(* IEC 61131-3 sources: 2026_Projet_YGO_ExcavatriceDragage/TOOLS/TEST_AUTO_CI/MOCKS, 9 files *)

(* ---- DEVICE_STATE.st ---- *)
(* =======================================================================
   📊 Type CODESYS système pour tests STruCpp
   ======================================================================= *)
TYPE DEVICE_STATE :
(
    UNKNOWN             := 0,
    STOPPED             := 1,
    CONFIG_ERROR        := 2,
    BUS_ERROR           := 3,
    DISABLED            := 4,
    INITIALIZING        := 5,
    RESET_ORIGIN        := 6,
    RESET_COMMUNICATION := 7,
    RESET_APPLICATION   := 8,
    RUNNING             := 9,
    LOGGER_ERROR        := 10
);
END_TYPE

(* ---- MOCK_GVL_IHM.st ---- *)
(* =======================================================================
   🧪 MOCK_GVL_IHM — Miroir TESTABLE de la GVL_IHM (harnais CI uniquement)
   ───────────────────────────────────────────────────────────────
   🎯 Pourquoi ce fichier existe (T371) :
      STruCpp v0.6.2 ne supporte PAS le namespace GVL de CODESYS. Une GVL
      `VAR_GLOBAL` déclare ses membres comme des variables GLOBALES PLATES :
      `GVL_IHM.Modes.Cmd.X` n'est donc pas résoluble, alors que c'est
      exactement ce que fait le code de production (CODESYS, où le nom de la
      GVL EST un espace de noms).
      Sonde compilateur (2026-09-21) : `VAR_GLOBAL Foo:INT;` + `GVL_T.Foo`
      -> "error: Undeclared variable 'GVL_T'" ; accès direct `Foo` -> OK ;
      `GVL_T` déclaré comme VARIABLE d'un STRUCT miroir -> OK.

   🔧 Principe : `GVL_IHM` est déclarée ici comme une VARIABLE GLOBALE d'un
      STRUCT MIROIR dont les membres sont la TRANSCRIPTION EXACTE de la liste
      de membres de `CODE/J_SUPERVISION/GVL_IHM.st`. Le code de production
      (`GVL_IHM.<membre>`) devient alors résoluble à l'identique.

   ⚠️ FICHIER DE TEST — JAMAIS compilé dans CODESYS, JAMAIS importé :
      il n'est référencé que par l'entrée `FB_TroubleshootingView` de
      `TOOLS/TEST_AUTO_CI/scripts/config/registry.yaml`.
   ⚠️ DETTE DÉCLARÉE : ce miroir peut dériver si `GVL_IHM.st` change. Une
      dérive produit une ERREUR DE COMPILATION du harnais (bruit), jamais un
      faux résultat silencieux. Toute évolution de `GVL_IHM.st` doit être
      répercutée ici.
   📄 Source de vérité transcrite : CODE/J_SUPERVISION/GVL_IHM.st:8-24
   ======================================================================= *)

TYPE ST_MockGvlIHM :
STRUCT
    M1TreuilRetenue    : ST_WinchHMI;               (* GVL_IHM.st:8  *)
    M2TreuilBenne      : ST_WinchBenneHMI;          (* GVL_IHM.st:9  — porte Bucket *)
    M1M2Sync           : ST_SyncHMI;                (* GVL_IHM.st:10 *)
    JOY1Joystick       : ST_JoystickHMI;            (* GVL_IHM.st:11 *)
    Modes              : ST_ModesHMI;               (* GVL_IHM.st:12 *)
    Emergency          : ST_EmergencyHMI;           (* GVL_IHM.st:13 *)
    M3Translation      : ST_TranslationHMI;         (* GVL_IHM.st:14 *)
    CycleSemiAuto      : ST_CycleHMI;               (* GVL_IHM.st:15 *)
    CycleMachineHoming : ST_CycleMachineHomingHMI;  (* GVL_IHM.st:16 *)
    Banner             : ST_HmiBanner;              (* GVL_IHM.st:17 *)
    Network            : ST_NetworkDiagHMI;         (* GVL_IHM.st:18 *)
    Commun             : ST_CommunHMI;              (* GVL_IHM.st:19 *)
    LocalIHM           : ST_LocalIHM;               (* GVL_IHM.st:20 *)
    IoHw               : ST_IoHw;                   (* GVL_IHM.st:21 *)
    HmiInitDone        : BOOL;                      (* GVL_IHM.st:22 *)
    Permits            : ST_PermitVisibilityHMI;    (* GVL_IHM.st:23 *)
    MaintenanceN2      : ST_MaintenanceN2HMI;       (* GVL_IHM.st:24 *)
END_STRUCT
END_TYPE

VAR_GLOBAL
    GVL_IHM : ST_MockGvlIHM;   // Miroir testable de la GVL de production (voir bandeau)
END_VAR

(* ---- MOCK_GVL_Troubleshooting.st ---- *)
(* =======================================================================
   🧪 MOCK_GVL_Troubleshooting — Miroir TESTABLE de la GVL_Troubleshooting
   ───────────────────────────────────────────────────────────────
   🎯 Pourquoi ce fichier existe (T371) : voir le bandeau détaillé de
      `TOOLS/TEST_AUTO_CI/MOCKS/MOCK_GVL_IHM.st` (même cause, même patron).
      En résumé : STruCpp v0.6.2 ne supporte pas le namespace GVL CODESYS ;
      `GVL_Troubleshooting.N_MotionM1.Step8_OutputInterlockOk` (écrit 469 fois
      par `FB_TroubleshootingView.st`) n'est résoluble que si `GVL_Troubleshooting`
      existe comme VARIABLE GLOBALE d'un STRUCT miroir — patron prouvé par sonde
      compilateur le 2026-09-21.

   ⚠️ FICHIER DE TEST — JAMAIS compilé dans CODESYS, JAMAIS importé :
      référencé uniquement par l'entrée `FB_TroubleshootingView` du registry CI.
   ⚠️ DETTE DÉCLARÉE : dérive possible si `GVL_Troubleshooting.st` change ->
      erreur de compilation du harnais (bruit), jamais un faux résultat silencieux.
   📄 Source de vérité transcrite : CODE/J_SUPERVISION/GVL_Troubleshooting.st
      (bloc VAR_GLOBAL, membres dans l'ordre du fichier source)
   ======================================================================= *)

TYPE ST_MockGvlTroubleshooting :
STRUCT
    A_ContexteMachineGlobal  : ST_ChainContextGlobal;   (* 0.  Contexte Global Machine *)
    B_Inputs                 : ST_HardwareImage;        (* 1.  Image complète des entrées *)
    C_Safety                 : ST_SafetyChecklist;      (* 2.  Chaîne de sécurité & réarmement AU *)
    D_Joystick               : ST_JoystickChecklist;    (* 3.  Bus CANopen & homme-mort joystick *)
    E_HomingM1               : ST_HomingChecklist;      (* 4.  Homing M1 *)
    F_HomingM2               : ST_HomingChecklist;      (* 5.  Homing M2 *)
    G_CycleSemiAuto          : ST_ChainCycleSemiAuto;   (* 6.  Séquenceur de cycle semi-auto *)
    H_LevageSynchroniseM1M2  : ST_ChainWinchSync;       (* 7.  Levage synchronisé M1+M2 *)
    I_LevageUnitaireM1       : ST_ChainWinch;           (* 8.  Levage unitaire M1 *)
    J_LevageUnitaireM2       : ST_ChainWinch;           (* 9.  Levage unitaire M2 *)
    K_BenneOuvertureFermeture: ST_ChainBucket;          (* 10. Ouverture / fermeture benne *)
    L_TranslationPontM3      : ST_ChainTranslation;     (* 11. Translation pont M3 *)
    N_MotionM1               : ST_MotionChecklist;      (* 13. Diagnostic mouvement M1 *)
    O_MotionM2               : ST_MotionChecklist;      (* 14. Diagnostic mouvement M2 *)
    P_MotionM3               : ST_MotionChecklist;      (* 15. Diagnostic mouvement M3 *)
    Q_TraceWinchM1           : ST_TraceWinch;           (* 16. Trace blocage M1 *)
    R_TraceWinchM2           : ST_TraceWinch;           (* 17. Trace blocage M2 *)
    S_TraceTranslation       : ST_TraceTranslation;     (* 18. Trace blocage M3 *)
    T_Permits                : ST_PermitVisibilityHMI;  (* Vue unique des permis *)
END_STRUCT
END_TYPE

VAR_GLOBAL
    GVL_Troubleshooting : ST_MockGvlTroubleshooting;   // Miroir testable de la GVL de production
END_VAR

(* ---- ST_fbJoystick_Cfg.st ---- *)
(* =======================================================================
   🧪 ST_fbJoystick_Cfg — Maquette STruCpp pour FB_SimBench
   -----------------------------------------------------------------------
   🎯 Rôle : satisfaire le champ ST_JoystickHMI.Cfg sans exercer FB_Joystick.
   📄 Portée : harnais STruCpp uniquement; le type production reste inchangé.
   ======================================================================= *)
TYPE ST_fbJoystick_Cfg :
STRUCT
END_STRUCT
END_TYPE

(* ---- ST_fbSim_Translation_ExtLink_Echo.st ---- *)
(* Test-only mirror of the retired external-M3 link payload.
   Production code no longer ships the OpenModelica link; FB_SimBench CI still
   requires its interface because MOCK_FB_Sim_Translation_ExtLink exposes it. *)
TYPE ST_fbSim_Translation_ExtLink_Echo :
STRUCT
    Mode                    : E_Mode;
    FBState                 : E_State;
    AxisBlockReason         : E_TranslationTraceBlockReason;
    MaintenanceTargetEnable : BOOL;
    MaintenanceZoneAccess   : BOOL;
    SafeStop                : BOOL;
    PowerCutOff             : BOOL;
    LimitSwitchTremie       : BOOL;
    LimitSwitchMaintenance  : BOOL;
    PositionReached         : BOOL;
    ActiveTremie            : BOOL;
    ActiveMaintenance       : BOOL;
    AtTremie                : BOOL;
    AtPV                    : BOOL;
    AtP2                    : BOOL;
    AtP1                    : BOOL;
    AtMaintenance           : BOOL;
    SensorWordIncoherent    : BOOL;
    EstimatedPos_M          : REAL;
    SafetyErrorId           : WORD;
END_STRUCT
END_TYPE

(* ---- FB_TestHarnessT417_M3.st ---- *)
(* T417 D2 — boucle fermee de preuve, composants de production composes dans l'ordre PRG02→PRG03/05→PRG06.
   Le cycle utilise ses entrees publiques. StepForceTgt ne sert qu'a fixer le point de depart AX14;
   les gestes, les transitions AX15A/B/C/18/2 et les demandes M3 restent emis par les vrais FB.
   M1/M2, benne, mode arbitre, IHM, reseaux et AU sont des faits de banc declares, pas couverts ici. *)
FUNCTION_BLOCK PUBLIC FB_TestHarnessT417_M3
VAR_INPUT
    Enable                  : BOOL;
    StepForceTgt            : INT := -1;
    JoystickLeft            : BOOL;
    JoystickRight           : BOOL;
    JoystickPush            : BOOL;
    JoystickPull            : BOOL;
    RepositionRequest       : BOOL;
    BenneDone               : BOOL;
    BenneIsOpen             : BOOL;
    SimM3Slope_Mps2         : REAL;
END_VAR
VAR_IN_OUT
    RawPosM1                : UDINT;
    RawPosM2                : UDINT;
END_VAR
VAR_OUTPUT
    CycleStep               : E_AutoCycleStep;
    CycleError              : BOOL;
    CycleReqStart            : BOOL;
    CyclePositionTgt          : INT;
    ArbitrationReqTremie      : BOOL;
    ArbitrationReqMaintenance : BOOL;
    ArbitrationRunRequest     : BOOL;
    TranslationSafetyError  : BOOL;
    TranslationMotionError  : BOOL;
    FinalInterlockError     : BOOL;
    M3ReqTremie              : BOOL;
    M3ReqMaintenance         : BOOL;
    M3DriveControlWord       : WORD;
    M3DriveFreqCmd_Hz        : REAL;
    M3DriveActualFreq_Hz     : REAL;
    M3BrakeReleaseRequest    : BOOL;
    M3BrakeFinalCmd          : BOOL;
    M3BrakeContactOpen       : BOOL;
    M3SensorsWord            : BYTE;
    M3AtTremie               : BOOL;
    M3AtP1                   : BOOL;
    M3PositionTrue_M         : REAL;
    M3PositionEstimated_M    : REAL;
    M3PositionError_M        : REAL;
    M3OvershootLast_M        : REAL;
    M3OvershootSensorId      : INT;
    P1ArrivalCaptured        : BOOL;
    P1ArrivalPosition_M       : REAL;
    P1ArrivalSensorsWord      : BYTE;
    P1ArrivalDriveControlWord : WORD;
    P1ArrivalFrequency_Hz     : REAL;
    P1ArrivalBrakeOpen        : BOOL;
    M3CartFree               : BOOL;
    M3FreeRollLast_M         : REAL;
END_VAR
VAR
    instCycle                : FB_CycleSemiAuto;
    instArbitration          : FB_TranslationCmdArbitrationM3;
    instSafety               : FB_Safety_Translation;
    instTranslation          : FB_Translation;
    instOutputInterlock      : FB_TranslationOutputInterlock;
    instPositionDecoder      : FB_Translation_PositionDecoder;
    instPositionEstimator    : FB_Translation_PositionEstimator;
    instSimBench             : FB_SimBench;
    TranslationCfg           : ST_fbTranslation_Cfg;
    Joystick                 : ST_AcquisitionJoystickQualified;
    ModesAuth                : ST_Modes_Autorisations;
    CycleTranslationRequest  : ST_ProgramTranslationRequest;
    ArbitrationIHM           : ST_fbTranslationCmdArbitration_IHM;
    ArbitrationContext       : ST_fbTranslationCmdArbitration_Context;
    ArbitrationCfg           : ST_fbTranslationCmdArbitration_Cfg;
    TargetCodeSel            : INT;
    SensorsWordPrev          : BYTE;
    SensorsWordChanged       : BOOL;
    PositionSensorTarget     : BOOL;
    AtTremieStable           : BOOL;
    AtPVStable               : BOOL;
    AtP2Stable               : BOOL;
    AtP1Stable               : BOOL;
    AtMaintenanceStable      : BOOL;
    AtPositionBootRestored   : BOOL;
    BootSensorsStable        : TON;
    SimReqTremieN1           : BOOL;
    SimReqMaintenanceN1      : BOOL;
    SimSpeedPctN1            : REAL;
    SimBrakeCmdN1            : BOOL;
    M3HeightInterlockOk      : BOOL;
    PermitTremie             : BOOL;
    PermitMaintenance        : BOOL;
    P1ArrivalCapturedLocal    : BOOL;
END_VAR

IF NOT Enable THEN
    CycleStep := E_AutoCycleStep.AX0_REPOS;
    RETURN;
END_IF;

(* La simulation est PRG02 : elle consomme les sorties finales mémorisées du scan N-1. *)
instSimBench(
    Enable := TRUE,
    OperatorSourceActive := TRUE,
    M3_ReqTremie := SimReqTremieN1,
    M3_ReqMaintenance := SimReqMaintenanceN1,
    M3_SpeedCmd_Pct := SimSpeedPctN1,
    M3_PosTremie_M := 0.0,
    M3_PosPV_M := 1.5,
    M3_PosP2_M := 3.5,
    M3_PosP1_M := 5.0,
    M3_PosMaintenance_M := 10.0,
    M3_OdometryGain := 0.02,
    M3_EstimatedPos_M := instPositionEstimator.PositionEstimatedM,
    M3_BrakeCmd := SimBrakeCmdN1,
    PowerKeepAlive_A := TRUE,
    PowerKeepAlive_B := TRUE,
    SimChainOkBit := TRUE,
    SimPhaseRotationOkBit := TRUE,
    SimM3SpeedFactor := 1.0,
    SimM3SensorIntermittenceActive := FALSE,
    SimM3SensorCamDropoutActive := FALSE,
    SimM3BrakePhysicalActive := TRUE,
    SimM3CartFreeActive := TRUE,
    SimM3LoadMassRatio := 0.5,
    SimM3RollingFriction_Mps2 := 0.1,
    SimM3Slope_Mps2 := SimM3Slope_Mps2,
    RawPosM1 := RawPosM1,
    RawPosM2 := RawPosM2
);

instPositionDecoder(
    SensorTremie := instSimBench.Translation.M3_PosTremie_DI,
    SensorPV := instSimBench.Translation.M3_PosPV_DI,
    SensorP2 := instSimBench.Translation.M3_PosPVP2_DI,
    SensorP1 := instSimBench.Translation.M3_PosP1_DI,
    SensorMaintenance := instSimBench.Translation.M3_PosMaintenance_DI
);

instPositionEstimator(
    Enable := TRUE,
    Reset := FALSE,
    DriveActualFreqHz := UINT_TO_REAL(instSimBench.Translation.M3_ActualFrequencyHz) / 100.0,
    ReqTremie := SimReqTremieN1,
    ReqMaintenance := SimReqMaintenanceN1,
    SensorMaintenance := instPositionDecoder.TranslationPosMaintenance,
    SensorP1 := instPositionDecoder.TranslationPosP1,
    SensorP2 := instPositionDecoder.TranslationPosP2,
    SensorPV := instPositionDecoder.TranslationPosPV,
    SensorTremie := instPositionDecoder.TranslationPosTremie,
    PosMaintenanceM := 10.0,
    PosP1M := 5.0,
    PosP2M := 3.5,
    PosPVM := 1.5,
    PosTremieM := 0.0,
    GainMetersPerHzSec := 0.02,
    PersistedPositionM := 0.0,
    PersistedInitialized := FALSE
);

SensorsWordChanged := instPositionDecoder.SensorsWord <> SensorsWordPrev;
BootSensorsStable(IN := NOT SimReqTremieN1 AND NOT SimReqMaintenanceN1, PT := T#500ms);
IF NOT AtPositionBootRestored AND BootSensorsStable.Q THEN
    CASE instPositionDecoder.SensorsWord OF
        2#11111: AtTremieStable := instPositionDecoder.TranslationPosTremie;
        2#01111: AtPVStable := instPositionDecoder.TranslationPosPV;
        2#00111: AtP2Stable := instPositionDecoder.TranslationPosP2;
        2#00011: AtP1Stable := instPositionDecoder.TranslationPosP1;
        2#00000: AtMaintenanceStable := instPositionDecoder.TranslationPosMaintenance;
    END_CASE;
    AtPositionBootRestored := TRUE;
ELSIF AtPositionBootRestored THEN
    IF instPositionDecoder.TranslationAtTremie THEN
        AtTremieStable := TRUE; AtPVStable := FALSE; AtP2Stable := FALSE; AtP1Stable := FALSE; AtMaintenanceStable := FALSE;
    ELSIF instPositionDecoder.TranslationAtPV THEN
        AtPVStable := TRUE; AtTremieStable := FALSE; AtP2Stable := FALSE; AtP1Stable := FALSE; AtMaintenanceStable := FALSE;
    ELSIF instPositionDecoder.TranslationAtP2 THEN
        AtP2Stable := TRUE; AtTremieStable := FALSE; AtPVStable := FALSE; AtP1Stable := FALSE; AtMaintenanceStable := FALSE;
    ELSIF instPositionDecoder.TranslationAtP1 THEN
        AtP1Stable := TRUE; AtTremieStable := FALSE; AtPVStable := FALSE; AtP2Stable := FALSE; AtMaintenanceStable := FALSE;
    ELSIF instPositionDecoder.TranslationAtMaintenance THEN
        AtMaintenanceStable := TRUE; AtTremieStable := FALSE; AtPVStable := FALSE; AtP2Stable := FALSE; AtP1Stable := FALSE;
    ELSIF SensorsWordChanged THEN
        AtPVStable := FALSE; AtP2Stable := FALSE; AtP1Stable := FALSE;
    END_IF;
    IF SimReqMaintenanceN1 THEN AtTremieStable := FALSE; END_IF;
    IF SimReqTremieN1 THEN AtMaintenanceStable := FALSE; END_IF;
END_IF;
SensorsWordPrev := instPositionDecoder.SensorsWord;

Joystick.AxisX.Enable := TRUE;
Joystick.AxisX.StartStop := JoystickLeft OR JoystickRight;
Joystick.AxisX.DirectionPositive := JoystickLeft;
Joystick.AxisX.DirectionNegative := JoystickRight;
Joystick.AxisX.AtNeutral := NOT JoystickLeft AND NOT JoystickRight;
Joystick.AxisX.Direction := SEL(JoystickLeft, SEL(JoystickRight, 0, -1), 1);
Joystick.AxisX.SpeedTgt := 100.0;
Joystick.AxisY.Enable := TRUE;
Joystick.AxisY.StartStop := JoystickPush OR JoystickPull;
Joystick.AxisY.DirectionPositive := JoystickPush;
Joystick.AxisY.DirectionNegative := JoystickPull;
Joystick.AxisY.AtNeutral := NOT JoystickPush AND NOT JoystickPull;
Joystick.AxisY.Direction := SEL(JoystickPush, SEL(JoystickPull, 0, -1), 1);
Joystick.AxisY.SpeedTgt := 100.0;
Joystick.DeadmanArmed := TRUE;
Joystick.AtNeutralXY := Joystick.AxisX.AtNeutral AND Joystick.AxisY.AtNeutral;
Joystick.Ready := TRUE;
ModesAuth.Mode := E_Mode.SEMI_AUTO;
ModesAuth.MaintenanceM3TargetEnable := FALSE;
M3HeightInterlockOk := TRUE; (* entree de banc declaree : M1/M2 au-dessus du seuil de PRG05 *)

instCycle(
    Enable := TRUE,
    PowerContactorEngaged := TRUE,
    EncoderFaultPresent := FALSE,
    Mode := E_Mode.SEMI_AUTO,
    JoystickDeflected := JoystickLeft OR JoystickRight OR JoystickPush OR JoystickPull,
    JoystickPush := JoystickPush,
    JoystickPull := JoystickPull,
    JoystickRight := JoystickRight,
    JoystickLeft := JoystickLeft,
    DeadmanArmed := TRUE,
    HeartbeatIhmOk := TRUE,
    SelTarget := 0,
    SetDepthM := -5.0,
    DepthStopMode := E_CycleDepthStopMode.KOBOLD_ONLY,
    WinchSyncError := FALSE,
    WinchSyncDeltaM := 0.0,
    M1_CablePosM := 5.0,
    M2_CablePosM := 5.0,
    M1_MeasuredSpeedMps := 0.0,
    M2_MeasuredSpeedMps := 0.0,
    M1_SpeedValid := TRUE,
    M2_SpeedValid := TRUE,
    M1_ContactorsReleased := TRUE,
    M2_ContactorsReleased := TRUE,
    M1_BrakeApplied := TRUE,
    M2_BrakeApplied := TRUE,
    SpeedMismatchThresholdMps := 0.0,
    SpeedMismatchTimeout := T#0ms,
    M1TopLimitReached := TRUE,
    M2TopLimitReached := TRUE,
    Translation_At_P1 := AtP1Stable,
    Translation_At_Tremie := AtTremieStable,
    Translation_At_Maintenance := AtMaintenanceStable,
    Translation_PosP1 := instPositionDecoder.TranslationPosP1,
    Translation_PosMaintenance := instPositionDecoder.TranslationPosMaintenance,
    Translation_Busy := ABS(instTranslation.RequestedDriveFreqHz) > 0.1,
    Translation_Done := instTranslation.TargetReached,
    Benne_Done := BenneDone,
    Benne_CloseReached := NOT BenneIsOpen,
    Benne_IsOpen := BenneIsOpen,
    Benne_IsClosed := NOT BenneIsOpen,
    Benne_IsRoughlyClosed := NOT BenneIsOpen,
    M1FinalAscentStartReady := TRUE,
    HomedM1 := TRUE,
    HomedM2 := TRUE,
    InitPositionOk := TRUE,
    WinchesAtTopWindow := TRUE,
    CfgDrainTime := T#0ms,
    RepositionRequest := RepositionRequest,
    StepForceTgt := StepForceTgt
);
CycleStep := instCycle.CycleStep;
CycleError := instCycle.Fault.Error;
CycleTranslationRequest := instCycle.TranslationCmd;
CycleReqStart := CycleTranslationRequest.ReqStart;
CyclePositionTgt := CycleTranslationRequest.PositionTgt;

ArbitrationContext.HeightInterlockOk := M3HeightInterlockOk;
ArbitrationCfg.MaxFreq_Hz := 50.0;
instArbitration(
    Enable := TRUE,
    Joystick := Joystick,
    Auth := ModesAuth,
    ReqTranslation := CycleTranslationRequest,
    IHM := ArbitrationIHM,
    TglJoystickMaster := FALSE,
    Context := ArbitrationContext,
    Cfg := ArbitrationCfg
);
ArbitrationReqTremie := instArbitration.ReqTremie;
ArbitrationReqMaintenance := instArbitration.ReqMaintenance;
ArbitrationRunRequest := instArbitration.RunRequest;
(* Le selecteur de cible est consommable au scan courant : retenir la derniere valeur non nulle. *)
IF instArbitration.SelTarget >= 1 AND instArbitration.SelTarget <= 4 THEN
    TargetCodeSel := instArbitration.SelTarget;
END_IF;
IF instArbitration.SelTarget = 0 THEN
    IF instArbitration.ReqTremie THEN
        TargetCodeSel := 1;
    ELSIF instArbitration.ReqMaintenance THEN
        TargetCodeSel := SEL(ModesAuth.MaintenanceM3TargetEnable, 3, 4);
    END_IF;
END_IF;
PositionSensorTarget := FALSE;
CASE TargetCodeSel OF
    1: PositionSensorTarget := AtTremieStable;
    2: PositionSensorTarget := AtP2Stable;
    3: PositionSensorTarget := AtP1Stable;
    4: PositionSensorTarget := AtMaintenanceStable;
END_CASE;

instSafety(
    Enable := TRUE,
    Reset := FALSE,
    PowerContactorEngaged := TRUE,
    Mode := E_Mode.SEMI_AUTO,
    JoystickOnline := TRUE,
    JoystickOperational := TRUE,
    HeartbeatIhmOk := TRUE,
    PhaseRotationOk := TRUE,
    BrakeThermalFeedback := FALSE,
    DriveOnline := TRUE,
    DriveOperational := TRUE,
    DriveStatusWord := instSimBench.Translation.M3_StatusWord,
    DriveActualFreqHz := UINT_TO_REAL(instSimBench.Translation.M3_ActualFrequencyHz) / 100.0,
    BrakeFeedback := instSimBench.Translation.M3_BrakeIsOpen_DI,
    BrakeCmd := instTranslation.BrakeReleaseRequest,
    RunRequest := instArbitration.RunRequest,
    ReqTremie := instArbitration.ReqTremie,
    ReqMaintenance := instArbitration.ReqMaintenance,
    LimitSwitchTremie := instPositionDecoder.LimitSwitchTremie,
    LimitSwitchMaintenance := instPositionDecoder.LimitSwitchMaintenance,
    SensorWordIncoherent := instPositionDecoder.Incoherent
);
PermitTremie := instSafety.TremieLimitClear AND NOT instSafety.SafeStop AND NOT instSafety.PowerCutOff;
PermitMaintenance := instSafety.MaintenanceLimitClear AND NOT instSafety.SafeStop AND NOT instSafety.PowerCutOff;

TranslationCfg.CfgRampAccelRate := 40.0;
TranslationCfg.CfgRampDecelNormalRate := 50.0;
TranslationCfg.CfgRampDecelFastRate := 100.0;
TranslationCfg.DriveFreqScaleMaxHz := 50.0;
TranslationCfg.ApproachSpeedTremieHz := 20.0;
TranslationCfg.ApproachSpeedMaintenanceHz := 20.0;
TranslationCfg.ApproachSpeedP1Hz := 20.0;
instTranslation(
    Enable := TRUE,
    Reset := FALSE,
    PowerContactorEngaged := TRUE,
    Mode := E_Mode.SEMI_AUTO,
    RunRequest := instArbitration.RunRequest,
    SafeStop := instSafety.SafeStop,
    ReqTremie := instArbitration.ReqTremie,
    ReqMaintenance := instArbitration.ReqMaintenance,
    SpeedTgt_Pct := instArbitration.SpeedPct,
    PositionSensorTarget := PositionSensorTarget,
    SlowdownSensorTremie := instPositionDecoder.TranslationPosPV,
    SlowdownSensorMaintenance := instPositionDecoder.TranslationPosP1,
    SlowdownSensorP1 := (NOT instPositionDecoder.TranslationPosP2) AND instPositionDecoder.TranslationPosP1,
    LimitSwitchTremie := instPositionDecoder.LimitSwitchTremie,
    LimitSwitchMaintenance := instPositionDecoder.LimitSwitchMaintenance,
    EffectivePermitM3_Tremie := PermitTremie,
    EffectivePermitM3_Maintenance := PermitMaintenance,
    DriveStatusWord := instSimBench.Translation.M3_StatusWord,
    DriveActualFreqHz := UINT_TO_REAL(instSimBench.Translation.M3_ActualFrequencyHz) / 100.0,
    BrakeFeedback := instSimBench.Translation.M3_BrakeIsOpen_DI,
    Cfg := TranslationCfg
);

instOutputInterlock(
    Enable := TRUE,
    Reset := FALSE,
    SafeStop := instSafety.SafeStop,
    PowerContactorEngaged := TRUE,
    EffectivePermitM3_Tremie := PermitTremie,
    EffectivePermitM3_Maintenance := PermitMaintenance,
    BrakeReleaseRequest := instTranslation.BrakeReleaseRequest,
    BrakeCommandOpenConfirmed := instTranslation.BrakeCommandOpenConfirmed,
    RequestedDriveControlWord := instTranslation.RequestedDriveControlWord,
    RequestedDriveFreqHz := instTranslation.RequestedDriveFreqHz
);

SimReqTremieN1 := instOutputInterlock.DriveControlWord = 1;
SimReqMaintenanceN1 := instOutputInterlock.DriveControlWord = 2;
SimSpeedPctN1 := (instOutputInterlock.DriveFreqCmd_Hz / 50.0) * 100.0;
SimBrakeCmdN1 := instOutputInterlock.BrakeCmd;

TranslationSafetyError := instSafety.Fault.Error;
TranslationMotionError := instTranslation.Fault.Error;
FinalInterlockError := instOutputInterlock.Fault.Error;
M3ReqTremie := SimReqTremieN1;
M3ReqMaintenance := SimReqMaintenanceN1;
M3DriveControlWord := instOutputInterlock.DriveControlWord;
M3DriveFreqCmd_Hz := instOutputInterlock.DriveFreqCmd_Hz;
M3DriveActualFreq_Hz := UINT_TO_REAL(instSimBench.Translation.M3_ActualFrequencyHz) / 100.0;
M3BrakeReleaseRequest := instTranslation.BrakeReleaseRequest;
M3BrakeFinalCmd := instOutputInterlock.BrakeCmd;
M3BrakeContactOpen := instSimBench.Translation.M3_BrakeIsOpen_DI;
M3SensorsWord := instPositionDecoder.SensorsWord;
M3AtTremie := AtTremieStable;
M3AtP1 := AtP1Stable;
M3PositionTrue_M := instSimBench.M3ObsPositionTrue_M;
M3PositionEstimated_M := instPositionEstimator.PositionEstimatedM;
M3PositionError_M := instSimBench.M3ObsPositionError_M;
M3OvershootLast_M := instSimBench.M3ObsOvershootLast_M;
M3OvershootSensorId := instSimBench.M3ObsOvershootSensorId;
IF (CycleStep = E_AutoCycleStep.AX18_DONE_SYNC) THEN
    P1ArrivalCapturedLocal := FALSE;
END_IF;
IF (CycleStep = E_AutoCycleStep.AX2_TRANSLATE_P1) AND AtP1Stable AND NOT P1ArrivalCapturedLocal THEN
    P1ArrivalCapturedLocal := TRUE;
    P1ArrivalCaptured := TRUE;
    P1ArrivalPosition_M := M3PositionTrue_M;
    P1ArrivalSensorsWord := M3SensorsWord;
    P1ArrivalDriveControlWord := M3DriveControlWord;
    P1ArrivalFrequency_Hz := M3DriveActualFreq_Hz;
    P1ArrivalBrakeOpen := M3BrakeContactOpen;
END_IF;
M3CartFree := instSimBench.M3ObsCartFree;
M3FreeRollLast_M := instSimBench.M3ObsFreeRollLast_M;
END_FUNCTION_BLOCK

(* ---- FB_TestLoopTranslation.st ---- *)
(* Harnais de test T417 : boucle fermee FB_Translation REEL (non modifie) + decodeur + FB_Sim_Translation.
   Un appel = un scan. Reproduit le cablage de PRG_05 (decodeur, ralentissements d approche, FdC bistable P1
   quand Maintenance est interdite, permis, jeton d arrivee P1). Non reproduit : FB_TranslationOutputInterlock
   (traite en transparent) et FB_Safety_Translation. Cible P1. Jamais compile dans le programme CODESYS. *)
FUNCTION_BLOCK FB_TestLoopTranslation
VAR_INPUT
    HoldRequest : BOOL;
END_VAR
VAR_OUTPUT
    Phase : INT;
    Overshoot_M : REAL;
    FreqAtCross_Hz : REAL;
    MaxCmdAfter_Hz : REAL;
    PositionTrue_M : REAL;
    CtrlWord : WORD;
    FreqReq_Hz : REAL;
    ActualFreq_Hz : REAL;
    AtP1Token : BOOL;
    SensorsWord : BYTE;
END_VAR
VAR
    tr : FB_Translation;
    sim : FB_Sim_Translation;
    dec : FB_Translation_PositionDecoder;
    cfg : ST_fbTranslation_Cfg;
    Initialized : BOOL;
    reqTremie : BOOL;
    reqMaint : BOOL;
    limTremieStable : BOOL;
    limMaintStable : BOOL;
    limMaintEff : BOOL;
    atP1 : BOOL;
    wordPrev : BYTE;
    wordChanged : BOOL;
    stopCount : INT;
    maxPos_M : REAL;
    crossed : BOOL;
END_VAR

IF NOT Initialized THEN
    Initialized := TRUE;
    cfg.CfgRampAccelRate := 40.0;
    cfg.CfgRampDecelNormalRate := 50.0;
    cfg.CfgRampDecelFastRate := 100.0;
    cfg.DriveFreqScaleMaxHz := 50.0;
    cfg.ApproachSpeedTremieHz := 20.0;
    cfg.ApproachSpeedMaintenanceHz := 20.0;
    cfg.ApproachSpeedP1Hz := 20.0;
    Phase := 0;
    reqTremie := TRUE;
END_IF;

dec(SensorTremie := sim.PosTremie, SensorPV := sim.PosPV, SensorP2 := sim.PosP2,
    SensorP1 := sim.PosP1, SensorMaintenance := sim.PosMaintenance);
limMaintEff := (NOT dec.TranslationPosP1) AND dec.TranslationPosMaintenance;
IF dec.LimitSwitchTremie THEN
    limTremieStable := TRUE;
ELSIF reqMaint THEN
    limTremieStable := FALSE;
END_IF;
IF limMaintEff THEN
    limMaintStable := TRUE;
ELSIF reqTremie THEN
    limMaintStable := FALSE;
END_IF;
wordChanged := (dec.SensorsWord <> wordPrev);
wordPrev := dec.SensorsWord;
IF dec.TranslationAtP1 THEN
    atP1 := TRUE;
ELSIF dec.TranslationAtP2 OR dec.TranslationAtPV OR dec.TranslationAtTremie OR dec.TranslationAtMaintenance OR wordChanged THEN
    atP1 := FALSE;
END_IF;

tr(Enable := TRUE, Reset := FALSE, PowerContactorEngaged := TRUE, RunRequest := TRUE, SafeStop := FALSE,
   ReqTremie := reqTremie, ReqMaintenance := reqMaint, SpeedTgt_Pct := 100.0,
   PositionSensorTarget := atP1 AND reqMaint,
   SlowdownSensorTremie := dec.TranslationPosPV,
   SlowdownSensorMaintenance := (NOT dec.TranslationPosP1) AND dec.TranslationPosMaintenance,
   SlowdownSensorP1 := (NOT dec.TranslationPosP2) AND dec.TranslationPosP1,
   LimitSwitchTremie := limTremieStable, LimitSwitchMaintenance := limMaintStable,
   EffectivePermitM3_Tremie := NOT limTremieStable, EffectivePermitM3_Maintenance := NOT limMaintStable,
   DriveStatusWord := 0, DriveActualFreqHz := sim.ActualFrequency_Hz,
   BrakeFeedback := sim.BrakeContactOpen, Cfg := cfg);
sim(Enable := TRUE,
    ReqTremie := (tr.RequestedDriveControlWord = 1), ReqMaintenance := (tr.RequestedDriveControlWord = 2),
    SpeedTgt_Pct := LIMIT(0.0, tr.RequestedDriveFreqHz / 50.0 * 100.0, 100.0),
    BrakeReleaseCmd := tr.BrakeReleaseRequest,
    LoadFrequencyDroopGain_Hz := 0.0, LoadReactionGain_Mps2 := 0.0);
PositionTrue_M := sim.PositionTrue_M;
CtrlWord := tr.RequestedDriveControlWord;
FreqReq_Hz := tr.RequestedDriveFreqHz;
ActualFreq_Hz := sim.ActualFrequency_Hz;
AtP1Token := atP1;
SensorsWord := dec.SensorsWord;

CASE Phase OF
    0:  (* jambe Tremie jusqu a 6 m : vitesse pleine atteinte hors zone d approche *)
        IF sim.PositionTrue_M < 6.0 THEN
            reqTremie := FALSE;
            Phase := 1;
            stopCount := 0;
        END_IF;
    1:  (* arret complet, frein ferme *)
        IF (sim.ActualFrequency_Hz < 0.5) AND (NOT sim.BrakeMechanicallyOpen) THEN
            stopCount := stopCount + 1;
        ELSE
            stopCount := 0;
        END_IF;
        IF stopCount > 30 THEN
            reqMaint := TRUE;
            Phase := 2;
        END_IF;
    2:  (* jambe Maintenance vers la cible P1 *)
        IF atP1 AND NOT HoldRequest THEN
            reqMaint := FALSE;
        END_IF;
        IF sim.PositionTrue_M > 20.0 THEN
            IF NOT crossed THEN
                crossed := TRUE;
                FreqAtCross_Hz := sim.ActualFrequency_Hz;
            END_IF;
            maxPos_M := MAX(maxPos_M, sim.PositionTrue_M);
            MaxCmdAfter_Hz := MAX(MaxCmdAfter_Hz, tr.RequestedDriveFreqHz);
        END_IF;
        IF crossed AND (sim.ActualFrequency_Hz < 0.5) AND (ABS(sim.VelocityTrue_Mps) < 0.01) THEN
            Phase := 3;
        END_IF;
END_CASE;
Overshoot_M := maxPos_M - 20.0;
END_FUNCTION_BLOCK

(* ---- HYSTERESIS.st ---- *)
(* =======================================================================
   📊 HYSTERESIS — Bibliothèque standard Util CODESYS (IN, HIGH, LOW -> OUT)
   ======================================================================= *)
FUNCTION_BLOCK FB_Hysteresis_Util
VAR_INPUT
    IN   : INT;
    HIGH : INT;
    LOW  : INT;
END_VAR
VAR_OUTPUT
    OUT  : BOOL := TRUE;
END_VAR

IF OUT THEN
    IF IN >= HIGH THEN
        OUT := FALSE;
    END_IF;
ELSE
    IF IN <= LOW THEN
        OUT := TRUE;
    END_IF;
END_IF;
END_FUNCTION_BLOCK

(* ---- MOCK_FB_Sim_Translation_ExtLink.st ---- *)
(* =======================================================================
   🧪 Mock FB_Sim_Translation_ExtLink — interface seule, sans socket UDP
   -----------------------------------------------------------------------
   Le FB réel (CODE/L_SIMULATION/FB_Sim_Translation_ExtLink.st) ouvre un socket
   loopback et initialise une structure par littéral : ni l'un ni l'autre ne
   compile sous STruCpp. Les tests FB_SimBench n'activent jamais la source
   externe M3 (SimM3OpenModelicaActive = FALSE) : seule l'interface compte.
   Interface recopiée à l'identique ; Enable=FALSE et TRUE -> lien jamais prêt.
   ======================================================================= *)
FUNCTION_BLOCK FB_Sim_Translation_ExtLink
VAR_INPUT
    Enable                  : BOOL;
    ReqTremie               : BOOL;
    ReqMaintenance          : BOOL;
    SetpointFrequencyHz     : WORD;
    BrakeReleaseCmd         : BOOL;
    PlcEcho                 : ST_fbSim_Translation_ExtLink_Echo;
END_VAR
VAR_OUTPUT
    Ready                   : BOOL;
    Translation             : ST_HwTranslation;
    LinkReady               : BOOL;
    LinkTimeout             : BOOL;
    LinkInvalid             : BOOL;
    LinkAge_Ms              : UDINT;
    TxCount                 : UDINT;
    RxCount                 : UDINT;
    RejectCount             : UDINT;
END_VAR

Ready := FALSE;
LinkReady := FALSE;
LinkTimeout := Enable;
LinkInvalid := Enable;
END_FUNCTION_BLOCK
